(* IEC 61131-3 sources: T4Exjobb/Sigma/Stations/MachineControl/MachineControl/Network/STDTimeSync, 1 file *)

(* ---- ONE_STDTimeSync_Table.st ---- *)
#define OBJECTS_CONFIG

#include <.\LoaderItf.h>
//Define part of class _SyncTimePLC
#define SyncTimeDate 60sec

FUNCTION GLOBAL TAB ONE_STDTimeSync
-1$UINT, 0$UINT,
2$UINT, 0$UINT,

5$UDINT,
TO_UDINT(4258542948), "_SIG_LSL_CMultimasterState", 1$UINT, 0$UINT, 1$UINT,
TO_UDINT(216306762), "_SyncTimePLC", 2$UINT, 0$UINT, 1$UINT,
TO_UDINT(3931827689), "_SysDateTime", 0$UINT, 7$UINT, 0$UINT,
TO_UDINT(3286875708), "_SysDateTime2", 0$UINT, 0$UINT, 1$UINT,
TO_UDINT(1903583397), "Ram", 1$UINT, 3$UINT, 1$UINT,

_NO_ATTR, TO_UDINT(3388907203), "_SIG_LSL_CMULTIMASTERSTATE1",

_NO_ATTR, TO_UDINT(1381574324), "SYNCTIMEPLC",

_NO_ATTR, TO_UDINT(985687168), "SYSDATETIMEPLC",

1$UINT, TO_UDINT(2994506371), "SYSDATETIMEPLC\_BASE\SUMMERTIME",

//Internal connections
0$UDINT,
1$UDINT,
TO_UDINT(2), "SummerTime", TO_UDINT(3),
0$UDINT,
3$UDINT,
TO_UDINT(1), "cOnline", TO_UDINT(0), "Terminal",
TO_UDINT(1), "cSetDate", TO_UDINT(2), "SysDate",
TO_UDINT(1), "cSetTime", TO_UDINT(2), "SysTime",

//Initialization values
0$UDINT,
1$UDINT,
TO_UDINT(2), "DoSummerTime", TO_UDINT(0),//|STDTimeSync.SysDateTimePLC.DoSummerTime;

//Symbolic initialization values
0$UDINT,
0$UDINT,

//Initialization of string values
0$UDINT,
0$UDINT,

//Configuration of tasks (RealTime, Cyclic, Background)
0$UDINT,
0$UDINT,

0$UDINT,
0$UDINT,

0$UDINT,
2$UDINT,
TO_UDINT(1), (10)$UDINT, 4194303$DINT, 	//SYNCTIMEPLC
TO_UDINT(2), (100)$UDINT, 4194303$DINT, 	//SYSDATETIMEPLC

//External connections
0$UDINT,
0$UDINT,

//Magic internal connections
0$UDINT,
0$UDINT,

//Configuration of timeslots of tasks (RealTime, Cyclic)
#ifdef __LSLLDR_TIMESLOTS__
0$UDINT,
0$UDINT,

0$UDINT,
0$UDINT,

#endif //__LSLLDR_TIMESLOTS__

//MultiMaster connections
#ifdef __LSLLDR_MULTIMASTER__
0$UDINT,
0$UDINT,
#endif //__LSLLDR_MULTIMASTER__

//Configuration for task ID (RealTime, CyclicTime)
#ifdef __LSLLDR_TASKID__
"\\\\TASKS2  "
0$UDINT,
0$UDINT,

0$UDINT,
0$UDINT,

0$UDINT,
2$UDINT,
(0)$UDINT, 	//SYNCTIMEPLC
(0)$UDINT, 	//SYSDATETIMEPLC

#endif //__LSLLDR_TASKID__

END_FUNCTION
